(* Logix 5000 project; controller WWTP_CLX vendor 1 type 14 code 54 rev 17.2; software revision 17.00; part 13 of 13 *)
(* tags used below, declared in another part *)
   I_AerTk_InflFlow : REAL;
   I_AerTk_InflFlow_IOFault : BOOL;
   I_AlumTk1Lv : ALIAS FOR WWTP_CLX_Rack01_Slot00_CNB:4:I.Ch0Data;
   I_AlumTk1Lv_IOFault : ALIAS FOR WWTP_CLX_Rack01_Slot00_CNB:4:I.Ch0Fault;
   LST1_CMPLX_CommFail : U_CommFail;
   PLC_Heartbeat : U_Heartbeat;
   PLC_Simulation : BOOL;   // Application running IN SIMULATION
   PLC_WallClock : U_WallClock;   // Wall Clock
   WWTP_AerTk_InflFlow : UD_Flow;   // Aeration Tank Influent Flow
   WWTP_AlumTk1Lv : P_AIn;   // Alum Tank #1 Level
   WWTP_CLX_Rack01_Slot00_Module : U_Module;
(* MainProgram, continued *)

ROUTINE A02_AnalogInputs   (* ladder *)
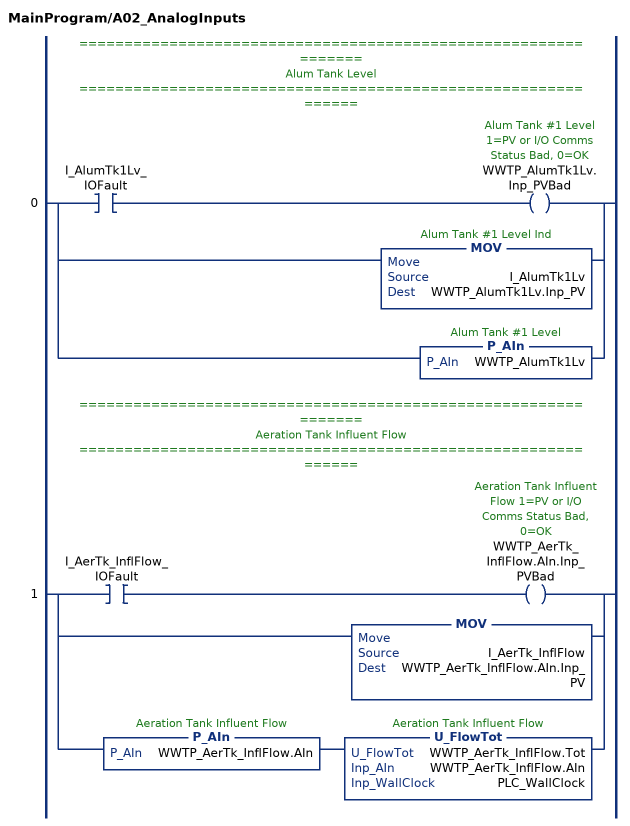
   // ===============================================================
   // Alum Tank Level
   // ==============================================================
   0: [XIC(I_AlumTk1Lv_IOFault) OTE(WWTP_AlumTk1Lv.Inp_PVBad) ,MOV(I_AlumTk1Lv,WWTP_AlumTk1Lv.Inp_PV) ,P_AIn(WWTP_AlumTk1Lv) ];
   // ===============================================================
   // Aeration Tank Influent Flow
   // ==============================================================
   1: [XIC(I_AerTk_InflFlow_IOFault) OTE(WWTP_AerTk_InflFlow.AIn.Inp_PVBad) ,MOV(I_AerTk_InflFlow,WWTP_AerTk_InflFlow.AIn.Inp_PV) ,P_AIn(WWTP_AerTk_InflFlow.AIn) U_FlowTot(WWTP_AerTk_InflFlow.Tot,WWTP_AerTk_InflFlow.AIn,PLC_WallClock) ];
END_ROUTINE

ROUTINE A03_DiscreteOutputs   (* ladder *)
   // ===============================================================
   // OUTPUT MAPPING
   // ===============================================================
   0: NOP();
END_ROUTINE

ROUTINE A04_AnalogOutputs   (* ladder *)
   // ===============================================================
   // OUTPUT MAPPING
   // ===============================================================
   0: NOP();
END_ROUTINE

ROUTINE Main   (* ladder *)
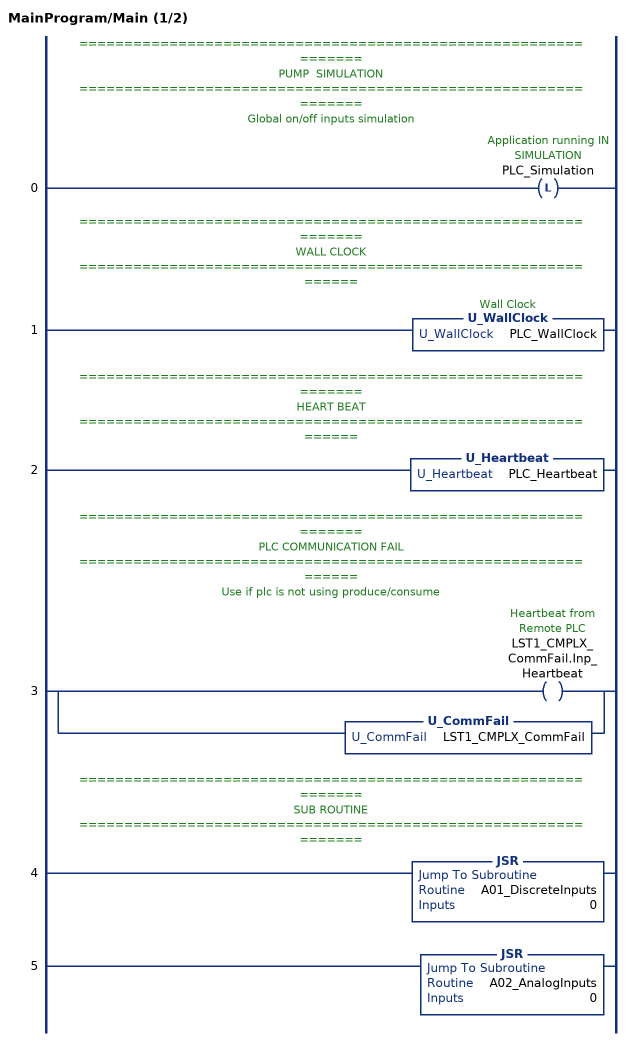
   // ===============================================================
   // PUMP  SIMULATION
   // ===============================================================
   // Global on/off inputs simulation
   0: OTL(PLC_Simulation);
   // ===============================================================
   // WALL CLOCK
   // ==============================================================
   1: U_WallClock(PLC_WallClock);
   // ===============================================================
   // HEART BEAT
   // ==============================================================
   2: U_Heartbeat(PLC_Heartbeat);
   // ===============================================================
   // PLC COMMUNICATION FAIL
   // ==============================================================
   // Use if plc is not using produce/consume
   3: [OTE(LST1_CMPLX_CommFail.Inp_Heartbeat) ,U_CommFail(LST1_CMPLX_CommFail) ];
   // ===============================================================
   // SUB ROUTINE
   // ===============================================================
   4: JSR(A01_DiscreteInputs,0);
   5: JSR(A02_AnalogInputs,0);
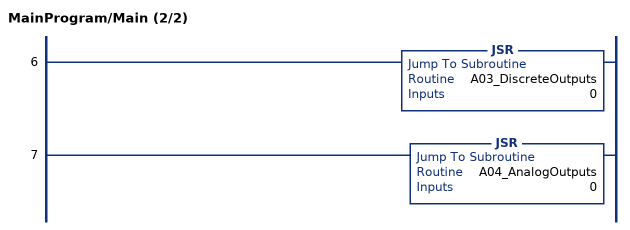
   6: JSR(A03_DiscreteOutputs,0);
   7: JSR(A04_AnalogOutputs,0);
END_ROUTINE
END_PROGRAM

PROGRAM MainTask   (* main routine MainProgram *)

ROUTINE MainProgram   (* ladder *)
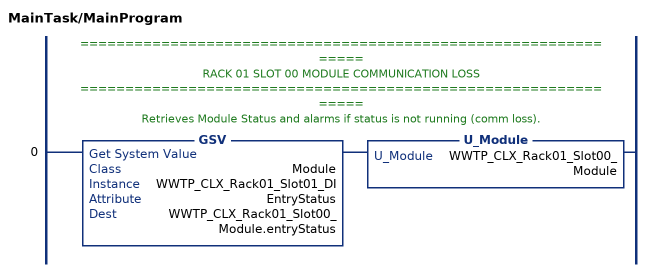
   // ===============================================================
   // RACK 01 SLOT 00 MODULE COMMUNICATION LOSS
   // ===============================================================
   // Retrieves Module Status and alarms if status is not running (comm loss).
   0: GSV(Module,WWTP_CLX_Rack01_Slot01_DI,EntryStatus,WWTP_CLX_Rack01_Slot00_Module.entryStatus)U_Module(WWTP_CLX_Rack01_Slot00_Module);
END_ROUTINE
END_PROGRAM
